(* IEC 61131-3 sources: rusty/tests/lit/multi/external_unit_linkage/chain/lib_c, 4 files *)

(* ---- base_of.st ---- *)
FUNCTION base_of : DINT
VAR_INPUT
    child : IChild;
END_VAR
VAR
    base : IBase;
END_VAR
    base := child;
    base_of := base.base_id() * 10 + child.child_id();
END_FUNCTION

(* ---- extra_of.st ---- *)
FUNCTION extra_of : DINT
VAR_INPUT
    extra : IExtra;
END_VAR
    extra_of := extra.extra();
END_FUNCTION

(* ---- shape_area.st ---- *)
FUNCTION shape_area : DINT
VAR_INPUT
    shape : IShape;
END_VAR
    shape_area := shape.area('km');
END_FUNCTION

(* ---- GrandChild.st ---- *)
FUNCTION_BLOCK GrandChild EXTENDS Concrete
    METHOD OVERRIDE area : DINT
    VAR_INPUT
        unit : STRING[10];
    END_VAR
        unit_seen := unit;
        area := 40;
    END_METHOD
END_FUNCTION_BLOCK
